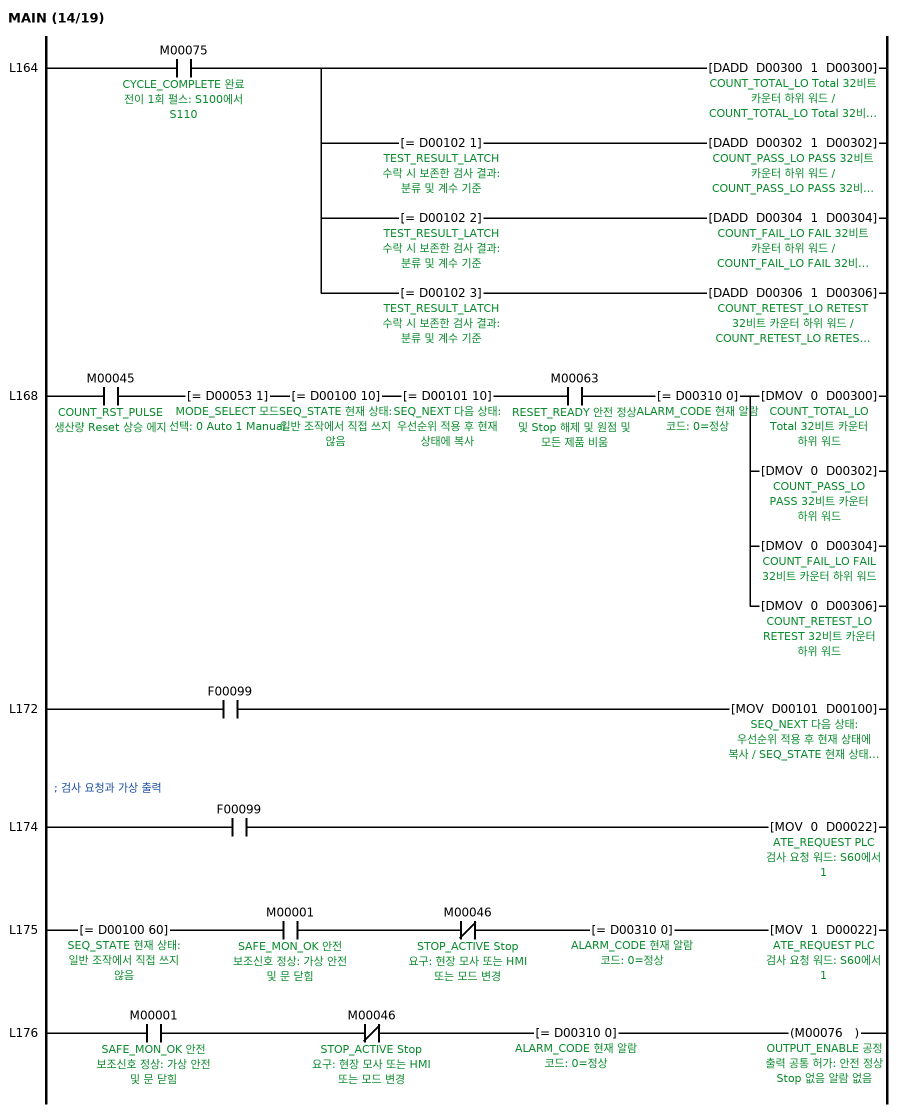
[picture p24: MAIN rungs L164-L176]
; L164
LOAD      M00075	// CYCLE_COMPLETE 완료 전이 1회 펄스: S100에서 S110
DADD      D00300 1 D00300	// COUNT_TOTAL_LO Total 32비트 카운터 하위 워드 / COUNT_TOTAL_LO Total 32비트 카운터 하위 워드
MPUSH
AND=      D00102 1	// TEST_RESULT_LATCH 수락 시 보존한 검사 결과: 분류 및 계수 기준
DADD      D00302 1 D00302	// COUNT_PASS_LO PASS 32비트 카운터 하위 워드 / COUNT_PASS_LO PASS 32비트 카운터 하위 워드
MLOAD
AND=      D00102 2	// TEST_RESULT_LATCH 수락 시 보존한 검사 결과: 분류 및 계수 기준
DADD      D00304 1 D00304	// COUNT_FAIL_LO FAIL 32비트 카운터 하위 워드 / COUNT_FAIL_LO FAIL 32비트 카운터 하위 워드
MPOP
AND=      D00102 3	// TEST_RESULT_LATCH 수락 시 보존한 검사 결과: 분류 및 계수 기준
DADD      D00306 1 D00306	// COUNT_RETEST_LO RETEST 32비트 카운터 하위 워드 / COUNT_RETEST_LO RETEST 32비트 카운터 하위 워드
; L168
LOAD      M00045	// COUNT_RST_PULSE 생산량 Reset 상승 에지
AND=      D00053 1	// MODE_SELECT 모드 선택: 0 Auto 1 Manual
AND=      D00100 10	// SEQ_STATE 현재 상태: 일반 조작에서 직접 쓰지 않음
AND=      D00101 10	// SEQ_NEXT 다음 상태: 우선순위 적용 후 현재 상태에 복사
AND       M00063	// RESET_READY 안전 정상 및 Stop 해제 및 원점 및 모든 제품 비움
AND=      D00310 0	// ALARM_CODE 현재 알람 코드: 0=정상
DMOV      0 D00300	// COUNT_TOTAL_LO Total 32비트 카운터 하위 워드
DMOV      0 D00302	// COUNT_PASS_LO PASS 32비트 카운터 하위 워드
DMOV      0 D00304	// COUNT_FAIL_LO FAIL 32비트 카운터 하위 워드
DMOV      0 D00306	// COUNT_RETEST_LO RETEST 32비트 카운터 하위 워드
; L172
LOAD      F00099
MOV       D00101 D00100	// SEQ_NEXT 다음 상태: 우선순위 적용 후 현재 상태에 복사 / SEQ_STATE 현재 상태: 일반 조작에서 직접 쓰지 않음
// 검사 요청과 가상 출력
; L174
LOAD      F00099
MOV       0 D00022	// ATE_REQUEST PLC 검사 요청 워드: S60에서 1
; L175
LOAD=     D00100 60	// SEQ_STATE 현재 상태: 일반 조작에서 직접 쓰지 않음
AND       M00001	// SAFE_MON_OK 안전 보조신호 정상: 가상 안전 및 문 닫힘
AND NOT   M00046	// STOP_ACTIVE Stop 요구: 현장 모사 또는 HMI 또는 모드 변경
AND=      D00310 0	// ALARM_CODE 현재 알람 코드: 0=정상
MOV       1 D00022	// ATE_REQUEST PLC 검사 요청 워드: S60에서 1
; L176
LOAD      M00001	// SAFE_MON_OK 안전 보조신호 정상: 가상 안전 및 문 닫힘
AND NOT   M00046	// STOP_ACTIVE Stop 요구: 현장 모사 또는 HMI 또는 모드 변경
AND=      D00310 0	// ALARM_CODE 현재 알람 코드: 0=정상
OUT       M00076	// OUTPUT_ENABLE 공정 출력 공통 허가: 안전 정상 Stop 없음 알람 없음

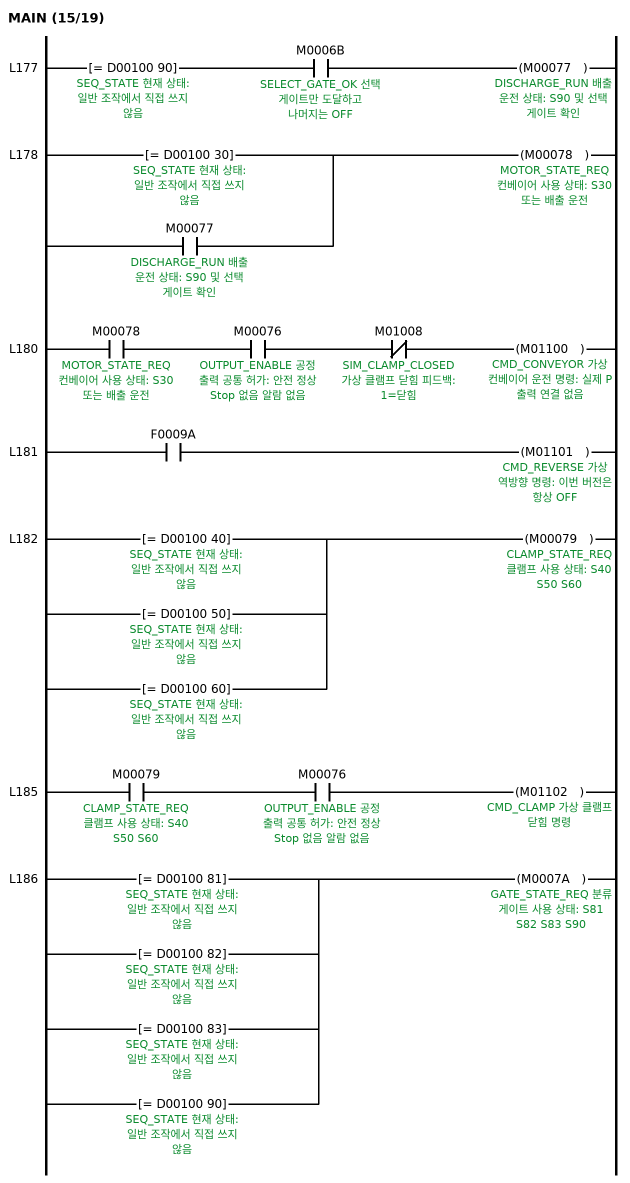
; L177
LOAD=     D00100 90	// SEQ_STATE 현재 상태: 일반 조작에서 직접 쓰지 않음
AND       M0006B	// SELECT_GATE_OK 선택 게이트만 도달하고 나머지는 OFF
OUT       M00077	// DISCHARGE_RUN 배출 운전 상태: S90 및 선택 게이트 확인
; L178
LOAD=     D00100 30	// SEQ_STATE 현재 상태: 일반 조작에서 직접 쓰지 않음
OR        M00077	// DISCHARGE_RUN 배출 운전 상태: S90 및 선택 게이트 확인
OUT       M00078	// MOTOR_STATE_REQ 컨베이어 사용 상태: S30 또는 배출 운전
; L180
LOAD      M00078	// MOTOR_STATE_REQ 컨베이어 사용 상태: S30 또는 배출 운전
AND       M00076	// OUTPUT_ENABLE 공정 출력 공통 허가: 안전 정상 Stop 없음 알람 없음
AND NOT   M01008	// SIM_CLAMP_CLOSED 가상 클램프 닫힘 피드백: 1=닫힘
OUT       M01100	// CMD_CONVEYOR 가상 컨베이어 운전 명령: 실제 P 출력 연결 없음
; L181
LOAD      F0009A
OUT       M01101	// CMD_REVERSE 가상 역방향 명령: 이번 버전은 항상 OFF
; L182
LOAD=     D00100 40	// SEQ_STATE 현재 상태: 일반 조작에서 직접 쓰지 않음
OR=       D00100 50	// SEQ_STATE 현재 상태: 일반 조작에서 직접 쓰지 않음
OR=       D00100 60	// SEQ_STATE 현재 상태: 일반 조작에서 직접 쓰지 않음
OUT       M00079	// CLAMP_STATE_REQ 클램프 사용 상태: S40 S50 S60
; L185
LOAD      M00079	// CLAMP_STATE_REQ 클램프 사용 상태: S40 S50 S60
AND       M00076	// OUTPUT_ENABLE 공정 출력 공통 허가: 안전 정상 Stop 없음 알람 없음
OUT       M01102	// CMD_CLAMP 가상 클램프 닫힘 명령
; L186
LOAD=     D00100 81	// SEQ_STATE 현재 상태: 일반 조작에서 직접 쓰지 않음
OR=       D00100 82	// SEQ_STATE 현재 상태: 일반 조작에서 직접 쓰지 않음
OR=       D00100 83	// SEQ_STATE 현재 상태: 일반 조작에서 직접 쓰지 않음
OR=       D00100 90	// SEQ_STATE 현재 상태: 일반 조작에서 직접 쓰지 않음
OUT       M0007A	// GATE_STATE_REQ 분류 게이트 사용 상태: S81 S82 S83 S90

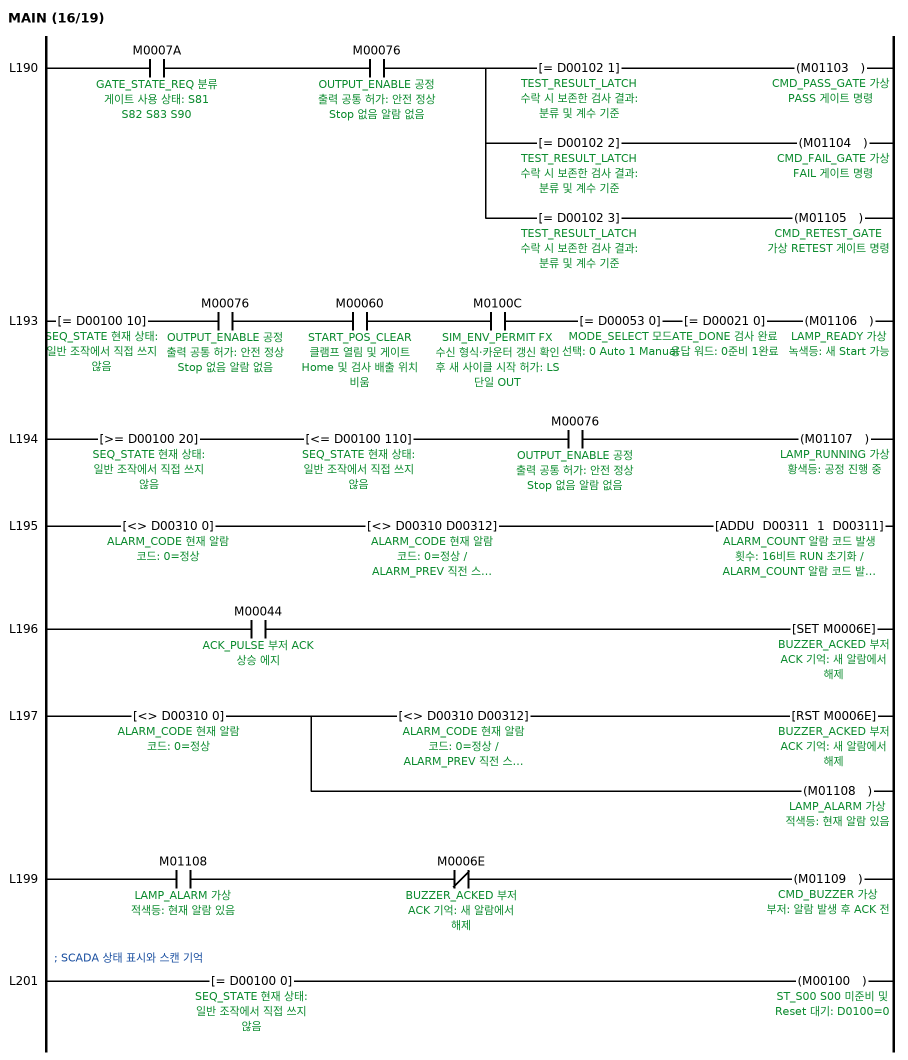
; L190
LOAD      M0007A	// GATE_STATE_REQ 분류 게이트 사용 상태: S81 S82 S83 S90
AND       M00076	// OUTPUT_ENABLE 공정 출력 공통 허가: 안전 정상 Stop 없음 알람 없음
MPUSH
AND=      D00102 1	// TEST_RESULT_LATCH 수락 시 보존한 검사 결과: 분류 및 계수 기준
OUT       M01103	// CMD_PASS_GATE 가상 PASS 게이트 명령
MLOAD
AND=      D00102 2	// TEST_RESULT_LATCH 수락 시 보존한 검사 결과: 분류 및 계수 기준
OUT       M01104	// CMD_FAIL_GATE 가상 FAIL 게이트 명령
MPOP
AND=      D00102 3	// TEST_RESULT_LATCH 수락 시 보존한 검사 결과: 분류 및 계수 기준
OUT       M01105	// CMD_RETEST_GATE 가상 RETEST 게이트 명령
; L193
LOAD=     D00100 10	// SEQ_STATE 현재 상태: 일반 조작에서 직접 쓰지 않음
AND       M00076	// OUTPUT_ENABLE 공정 출력 공통 허가: 안전 정상 Stop 없음 알람 없음
AND       M00060	// START_POS_CLEAR 클램프 열림 및 게이트 Home 및 검사 배출 위치 비움
AND       M0100C	// SIM_ENV_PERMIT FX 수신 형식·카운터 갱신 확인 후 새 사이클 시작 허가: LS 단일 OUT
AND=      D00053 0	// MODE_SELECT 모드 선택: 0 Auto 1 Manual
AND=      D00021 0	// ATE_DONE 검사 완료 응답 워드: 0준비 1완료
OUT       M01106	// LAMP_READY 가상 녹색등: 새 Start 가능
; L194
LOAD>=    D00100 20	// SEQ_STATE 현재 상태: 일반 조작에서 직접 쓰지 않음
AND<=     D00100 110	// SEQ_STATE 현재 상태: 일반 조작에서 직접 쓰지 않음
AND       M00076	// OUTPUT_ENABLE 공정 출력 공통 허가: 안전 정상 Stop 없음 알람 없음
OUT       M01107	// LAMP_RUNNING 가상 황색등: 공정 진행 중
; L195
LOAD<>    D00310 0	// ALARM_CODE 현재 알람 코드: 0=정상
AND<>     D00310 D00312	// ALARM_CODE 현재 알람 코드: 0=정상 / ALARM_PREV 직전 스캔 알람 코드: 새 알람 판정용
ADDU      D00311 1 D00311	// ALARM_COUNT 알람 코드 발생 횟수: 16비트 RUN 초기화 / ALARM_COUNT 알람 코드 발생 횟수: 16비트 RUN 초기화
; L196
LOAD      M00044	// ACK_PULSE 부저 ACK 상승 에지
SET       M0006E	// BUZZER_ACKED 부저 ACK 기억: 새 알람에서 해제
; L197
LOAD<>    D00310 0	// ALARM_CODE 현재 알람 코드: 0=정상
MPUSH
AND<>     D00310 D00312	// ALARM_CODE 현재 알람 코드: 0=정상 / ALARM_PREV 직전 스캔 알람 코드: 새 알람 판정용
RST       M0006E	// BUZZER_ACKED 부저 ACK 기억: 새 알람에서 해제
MPOP
OUT       M01108	// LAMP_ALARM 가상 적색등: 현재 알람 있음
; L199
LOAD      M01108	// LAMP_ALARM 가상 적색등: 현재 알람 있음
AND NOT   M0006E	// BUZZER_ACKED 부저 ACK 기억: 새 알람에서 해제
OUT       M01109	// CMD_BUZZER 가상 부저: 알람 발생 후 ACK 전
// SCADA 상태 표시와 스캔 기억
; L201
LOAD=     D00100 0	// SEQ_STATE 현재 상태: 일반 조작에서 직접 쓰지 않음
OUT       M00100	// ST_S00 S00 미준비 및 Reset 대기: D0100=0

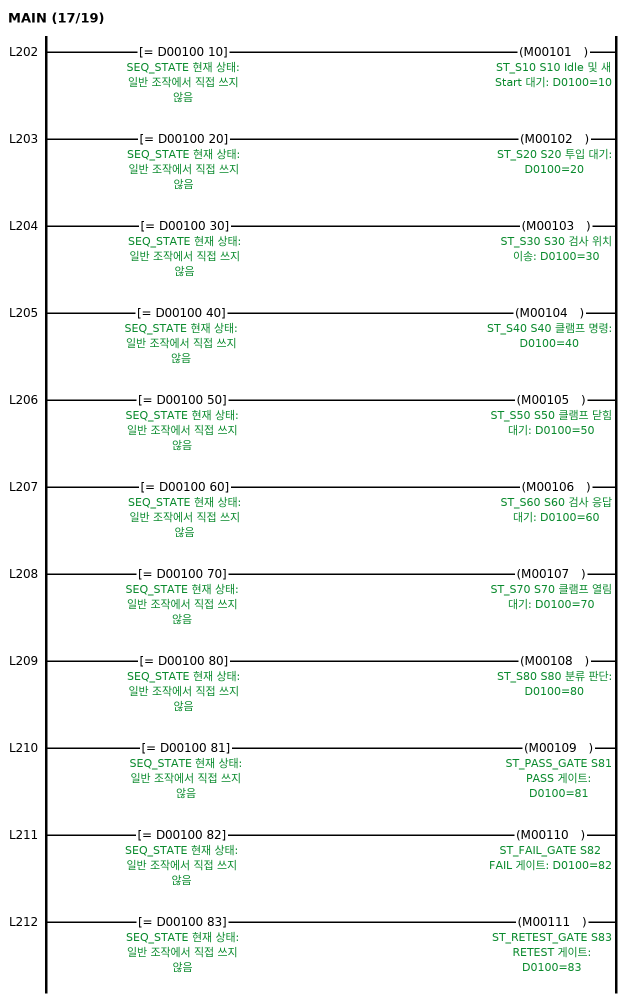
; L202
LOAD=     D00100 10	// SEQ_STATE 현재 상태: 일반 조작에서 직접 쓰지 않음
OUT       M00101	// ST_S10 S10 Idle 및 새 Start 대기: D0100=10
; L203
LOAD=     D00100 20	// SEQ_STATE 현재 상태: 일반 조작에서 직접 쓰지 않음
OUT       M00102	// ST_S20 S20 투입 대기: D0100=20
; L204
LOAD=     D00100 30	// SEQ_STATE 현재 상태: 일반 조작에서 직접 쓰지 않음
OUT       M00103	// ST_S30 S30 검사 위치 이송: D0100=30
; L205
LOAD=     D00100 40	// SEQ_STATE 현재 상태: 일반 조작에서 직접 쓰지 않음
OUT       M00104	// ST_S40 S40 클램프 명령: D0100=40
; L206
LOAD=     D00100 50	// SEQ_STATE 현재 상태: 일반 조작에서 직접 쓰지 않음
OUT       M00105	// ST_S50 S50 클램프 닫힘 대기: D0100=50
; L207
LOAD=     D00100 60	// SEQ_STATE 현재 상태: 일반 조작에서 직접 쓰지 않음
OUT       M00106	// ST_S60 S60 검사 응답 대기: D0100=60
; L208
LOAD=     D00100 70	// SEQ_STATE 현재 상태: 일반 조작에서 직접 쓰지 않음
OUT       M00107	// ST_S70 S70 클램프 열림 대기: D0100=70
; L209
LOAD=     D00100 80	// SEQ_STATE 현재 상태: 일반 조작에서 직접 쓰지 않음
OUT       M00108	// ST_S80 S80 분류 판단: D0100=80
; L210
LOAD=     D00100 81	// SEQ_STATE 현재 상태: 일반 조작에서 직접 쓰지 않음
OUT       M00109	// ST_PASS_GATE S81 PASS 게이트: D0100=81
; L211
LOAD=     D00100 82	// SEQ_STATE 현재 상태: 일반 조작에서 직접 쓰지 않음
OUT       M00110	// ST_FAIL_GATE S82 FAIL 게이트: D0100=82
; L212
LOAD=     D00100 83	// SEQ_STATE 현재 상태: 일반 조작에서 직접 쓰지 않음
OUT       M00111	// ST_RETEST_GATE S83 RETEST 게이트: D0100=83

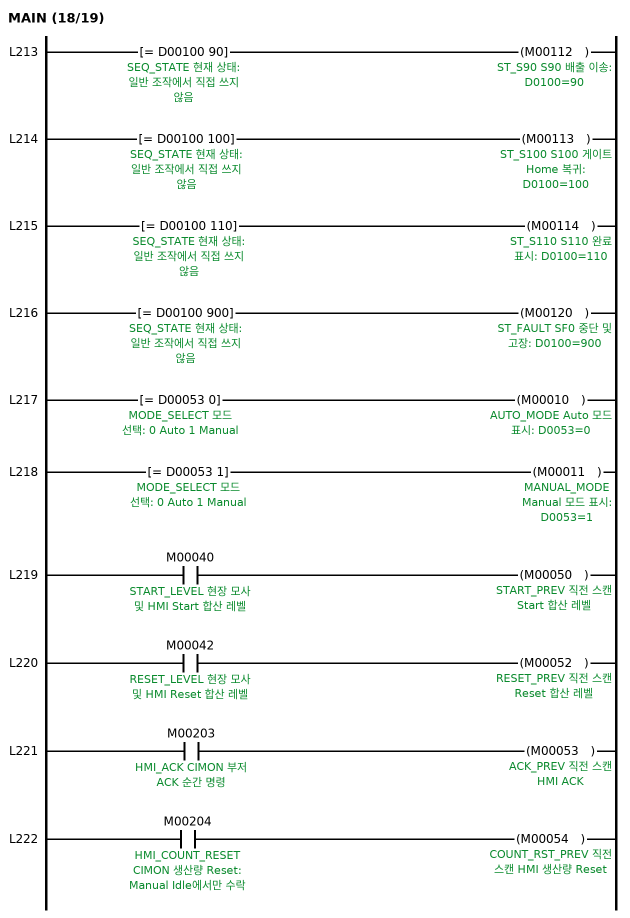
; L213
LOAD=     D00100 90	// SEQ_STATE 현재 상태: 일반 조작에서 직접 쓰지 않음
OUT       M00112	// ST_S90 S90 배출 이송: D0100=90
; L214
LOAD=     D00100 100	// SEQ_STATE 현재 상태: 일반 조작에서 직접 쓰지 않음
OUT       M00113	// ST_S100 S100 게이트 Home 복귀: D0100=100
; L215
LOAD=     D00100 110	// SEQ_STATE 현재 상태: 일반 조작에서 직접 쓰지 않음
OUT       M00114	// ST_S110 S110 완료 표시: D0100=110
; L216
LOAD=     D00100 900	// SEQ_STATE 현재 상태: 일반 조작에서 직접 쓰지 않음
OUT       M00120	// ST_FAULT SF0 중단 및 고장: D0100=900
; L217
LOAD=     D00053 0	// MODE_SELECT 모드 선택: 0 Auto 1 Manual
OUT       M00010	// AUTO_MODE Auto 모드 표시: D0053=0
; L218
LOAD=     D00053 1	// MODE_SELECT 모드 선택: 0 Auto 1 Manual
OUT       M00011	// MANUAL_MODE Manual 모드 표시: D0053=1
; L219
LOAD      M00040	// START_LEVEL 현장 모사 및 HMI Start 합산 레벨
OUT       M00050	// START_PREV 직전 스캔 Start 합산 레벨
; L220
LOAD      M00042	// RESET_LEVEL 현장 모사 및 HMI Reset 합산 레벨
OUT       M00052	// RESET_PREV 직전 스캔 Reset 합산 레벨
; L221
LOAD      M00203	// HMI_ACK CIMON 부저 ACK 순간 명령
OUT       M00053	// ACK_PREV 직전 스캔 HMI ACK
; L222
LOAD      M00204	// HMI_COUNT_RESET CIMON 생산량 Reset: Manual Idle에서만 수락
OUT       M00054	// COUNT_RST_PREV 직전 스캔 HMI 생산량 Reset

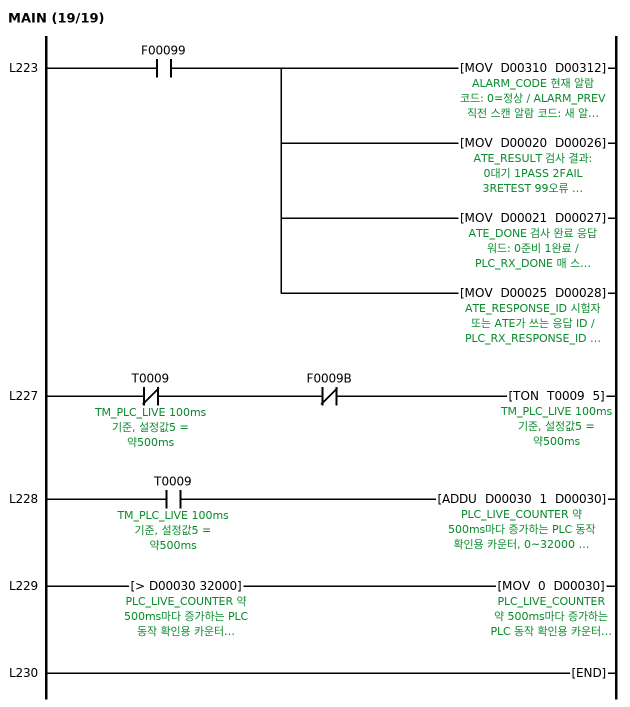
; L223
LOAD      F00099
MOV       D00310 D00312	// ALARM_CODE 현재 알람 코드: 0=정상 / ALARM_PREV 직전 스캔 알람 코드: 새 알람 판정용
MOV       D00020 D00026	// ATE_RESULT 검사 결과: 0대기 1PASS 2FAIL 3RETEST 99오류 / PLC_RX_RESULT 매 스캔 D00020을 복사한 실제 수신 결과
MOV       D00021 D00027	// ATE_DONE 검사 완료 응답 워드: 0준비 1완료 / PLC_RX_DONE 매 스캔 D00021을 복사한 실제 DONE
MOV       D00025 D00028	// ATE_RESPONSE_ID 시험자 또는 ATE가 쓰는 응답 ID / PLC_RX_RESPONSE_ID 매 스캔 D00025를 복사한 실제 응답 ID
; L227
LOAD NOT  T0009	// TM_PLC_LIVE 100ms 기준, 설정값5 = 약500ms
AND NOT   F0009B
TON       T0009 5	// TM_PLC_LIVE 100ms 기준, 설정값5 = 약500ms
; L228
LOAD      T0009	// TM_PLC_LIVE 100ms 기준, 설정값5 = 약500ms
ADDU      D00030 1 D00030	// PLC_LIVE_COUNTER 약 500ms마다 증가하는 PLC 동작 확인용 카운터, 0~32000 / PLC_LIVE_COUNTER 약 500ms마다 증가하는 PLC 동작 확인용 카운터, 0~32000
; L229
LOAD>     D00030 32000	// PLC_LIVE_COUNTER 약 500ms마다 증가하는 PLC 동작 확인용 카운터, 0~32000
MOV       0 D00030	// PLC_LIVE_COUNTER 약 500ms마다 증가하는 PLC 동작 확인용 카운터, 0~32000
; L230
END

VARIABLES AND COMMENTS (devices not used above)
D00023	WORD	ATE_HEARTBEAT_RSVD // 예약: ATE 하트비트 감시 미구현
D00305	WORD	COUNT_FAIL_HI // FAIL 32비트 카운터 상위 워드
D00303	WORD	COUNT_PASS_HI // PASS 32비트 카운터 상위 워드
D00307	WORD	COUNT_RETEST_HI // RETEST 32비트 카운터 상위 워드
D00301	WORD	COUNT_TOTAL_HI // Total 32비트 카운터 상위 워드
D00405	WORD	FX_ENV_CODE_REM // DIV 나머지. 다른 변수 배정 금지 / LS
D00408	WORD	FX_ENV_HB_REM // DIV 나머지. 다른 변수 배정 금지 / LS
D00206	WORD	PT_COMM_RSVD // 예약: 통신 시간 설정 미구현
T0007	BIT/WORD	TM_COMM_RSVD // 예약: 통신 감시 타이머 미구현